Fanuc KAREL source: KA00182.KL

PROGRAM KA00182
%NOLOCKGROUP
VAR
  SRC: ARRAY[4] OF BYTE
  DST: ARRAY[4] OF REAL
BEGIN
  DST = SRC
END KA00182
